(* IEC 61131-3 sources: kns-port-domestic/tools/plcopen/tests/fixtures/constructs/src/POUs/PRG_Main, 2 files *)

(* ---- PRG_Main.decl.st ---- *)
// Назначение: точка входа — вызывает все объекты примера
// Автор:      <ИМЯ ФАМИЛИЯ>
// Версия:     0.1.0
// Документ:   docs/plcopen.md
PROGRAM PRG_Main
VAR
    fbMotor : FB_Motor;
    itfDevice : I_Device;
    itfReset : I_Resettable;
    fbCounter : FB_Counter;
    stCmd : ST_MotorCmd;
    stSts : ST_MotorSts;
    stDerived : ST_Derived;
    uRaw : U_Raw;
    ePercent : T_Percent := 50;
    sName : T_Name := 'pump';
    eColor : E_Color := E_Color.Green;
    arBuf : ARRAY[0..2] OF REAL := [3(1.0)];
    rOut : REAL;
    lrSum : LREAL;
    pValue : POINTER TO REAL;
    refValue : REFERENCE TO REAL;
    iStep : INT;
    xOk : BOOL;
END_VAR

(* ---- PRG_Main.impl.st ---- *)
(* вызовы всех объектов примера *)
itfDevice := fbMotor;
itfReset := fbMotor;
fbMotor(stCmd := stCmd);
IF itfDevice <> 0 THEN
    itfDevice.Mode := E_Mode.Auto;
    xOk := itfDevice.Fault;
END_IF
itfReset.Reset(xForce := TRUE);
fbCounter(xIn := GVL_Io.xDiStart, stCmd := GVL_Io.astCmd[GVL_Io.IO_CHANNELS - 1]);
GVL_Io.xDoRun := fbMotor.xRun;
stSts.xRun := fbMotor.xRun;
stSts.uiStarts := fbMotor.Starts;
rOut := F_Clamp(rValue := INT_TO_REAL(GVL_Io.iAiLevel), rMin := 0.0, rMax := 100.0);
lrSum := F_Sum(arValues := arBuf);
pValue := ADR(rOut);
refValue REF= rOut;
IF __ISVALIDREF(refValue) THEN
    refValue := refValue + GVL_Const.RATE_LIMIT;
END_IF
uRaw.wWord := 16#1234;
stDerived.tDelay := T#1S;
CASE iStep OF
    0:
        iStep := 1;
    1, 2:
        iStep := iStep + 1;
ELSE
    iStep := 0;
END_CASE
WHILE iStep > 10 DO
    iStep := iStep - 1;
END_WHILE
REPEAT
    iStep := iStep + 0;
UNTIL TRUE
END_REPEAT
GVL_Io.udiRunHours := GVL_Io.udiRunHours + fbCounter.udiCount;
PersistentVars.udiStartsTotal := PersistentVars.udiStartsTotal + fbMotor.Starts;
sName := GVL_Const.TEXT_OK;
eColor := E_Color.Blue;
ePercent := 75;
PRG_Aux();
